(*
SPDX-License-Identifier: MIT
License: https://opensource.org/license/mit
*)

(*!
<summary>Runs an owned group containing a test controlled by its deadline.</summary>
<description>
Owns persistent root instances and fixed child storage. Use from one task without reentry.
Children borrows the same array for the instance lifetime. Root parents remain zero.
</description>
*)

{attribute 'no_assign'}
{attribute 'no_explicit_call' := 'do not call this function block directly'}
FUNCTION_BLOCK DeadlineTestRunner EXTENDS TOF_Testing.TestRunner<1>
VAR_STAT
	//! <summary>Class name shared by instances of this concrete runner.</summary>
	{attribute 'hide'}
	_ClassName : STRING := __POUNAME();
END_VAR
VAR
	{attribute 'hide'}
	{attribute 'init_namespace'}
	_NamespaceName : STRING;
END_VAR
VAR_OUTPUT
	//! <summary>Owned root element used by this runner.</summary>
	DeadlineGroup : DeadlineTestGroup(name := "Deadline group", parent := 0);
END_VAR
VAR
	_Children : ARRAY [0.._ChildCount - 1] OF TOF_Testing.ITestElement :=
	[
		DeadlineGroup
	];
END_VAR

(*!
<summary>Borrows the concrete class name; callers must not modify the returned storage.</summary>
*)
{attribute 'monitoring' := 'call'}
PROPERTY ClassName : REFERENCE TO STRING
GET
ClassName REF= _ClassName;
END_GET
END_PROPERTY

(*!
<summary>Borrows the concrete namespace name for the instance lifetime; callers must not modify it.</summary>
*)
{attribute 'monitoring' := 'call'}
PROPERTY NamespaceName : REFERENCE TO STRING
GET
NamespaceName REF= _NamespaceName;
END_GET
END_PROPERTY

(*!
<summary>Reports the complete concrete instance size.</summary>
*)
{attribute 'monitoring' := 'call'}
PROPERTY SelfSize : ULINT
GET
SelfSize := XSIZEOF(THIS^);
END_GET
END_PROPERTY

(*!
<summary>Borrows the unchanged persistent root array; application code must not modify it.</summary>
*)
{attribute 'monitoring' := 'call'}
PROPERTY Children : REFERENCE TO ARRAY [0.._ChildCount - 1] OF TOF_Testing.ITestElement
GET
Children REF= _Children;
END_GET
END_PROPERTY

END_FUNCTION_BLOCK

(* stored: Version 1.1.0.1
   POU DeadlineTestRunner: Id {fb3417fc-c7d7-49c0-9797-daaedb09d8da}, SpecialFunc None
   Property ClassName: Id {249f6ce6-5832-46e5-9846-bb56ba6d3a5b}
   Get Get: Id {61b618e2-3946-495e-8c49-317e16d118e2}
   Property NamespaceName: Id {03b5e773-9158-46ac-845e-a8fe7706ffe8}
   Get Get: Id {04fd0d5c-565d-44a9-9d7d-94cd460e5378}
   Property SelfSize: Id {433ddae9-205f-4cbe-9fda-859c87a75068}
   Get Get: Id {60eaf698-1c51-4990-a421-662145b9e8c6}
   Property Children: Id {84a66152-f772-49d0-a9cb-2efa3af14090}
   Get Get: Id {fbb127af-d19e-4986-b8bf-174950d64842} *)
